(* IEC 61131-3 sources: test/Network/Pump, 1 file *)

(* ---- ONE_Pump_Table.st ---- *)
#define OBJECTS_CONFIG

//Define part of class pumpControl
#define test 1

FUNCTION GLOBAL TAB ONE_Pump
-1$UINT, 0$UINT,
0$UINT, 0$UINT,

1$UDINT,
TO_UDINT(2030910333), "pumpControl", 0$UINT, 0$UINT, 2$UINT,

_NO_ATTR, TO_UDINT(2903633677), "PUMPCONTROL1",
_NO_ATTR, TO_UDINT(874036919), "PUMPCONTROL2",

//Internal connections
0$UDINT,
0$UDINT,
0$UDINT,
0$UDINT,

//Initialization values
0$UDINT,
6$UDINT,
TO_UDINT(0), "MaxBorder", TO_UDINT(800),//|Pump.pumpControl1.MaxBorder;
TO_UDINT(0), "Pump", TO_UDINT(0),//|Pump.pumpControl1.Pump;
TO_UDINT(0), "ActFillLevel", TO_UDINT(0),//|Pump.pumpControl1.ActFillLevel;
TO_UDINT(1), "MaxBorder", TO_UDINT(800),//|Pump.pumpControl2.MaxBorder;
TO_UDINT(1), "Pump", TO_UDINT(0),//|Pump.pumpControl2.Pump;
TO_UDINT(1), "ActFillLevel", TO_UDINT(0),//|Pump.pumpControl2.ActFillLevel;

//Symbolic initialization values
0$UDINT,
0$UDINT,

//Initialization of string values
0$UDINT,
0$UDINT,

//Configuration of tasks (RealTime, Cyclic, Background)
0$UDINT,
0$UDINT,

0$UDINT,
2$UDINT,
TO_UDINT(0), (10)$UDINT, 4194303$DINT, 	//PUMPCONTROL1
TO_UDINT(1), (10)$UDINT, 4194303$DINT, 	//PUMPCONTROL2

0$UDINT,
0$UDINT,

//External connections
0$UDINT,
3$UDINT,
TO_UDINT(0), "ActFillLevel", C_TRY, TO_UDINT(1457099445), "AI0431","AI2",
TO_UDINT(0), "test2", C_TRY, TO_UDINT(4130059223), "SDM0811","Safe_Input1",
TO_UDINT(0), "test1", C_TRY, TO_UDINT(4130059223), "SDM0811","Safe_Input2",

//Magic internal connections
0$UDINT,
0$UDINT,

//Configuration of timeslots of tasks (RealTime, Cyclic)
#ifdef __LSLLDR_TIMESLOTS__
0$UDINT,
0$UDINT,

0$UDINT,
0$UDINT,

#endif //__LSLLDR_TIMESLOTS__

//MultiMaster connections
#ifdef __LSLLDR_MULTIMASTER__
0$UDINT,
0$UDINT,
#endif //__LSLLDR_MULTIMASTER__

//Configuration for task ID (RealTime, CyclicTime)
#ifdef __LSLLDR_TASKID__
"\\\\TASKS2  "
0$UDINT,
0$UDINT,

0$UDINT,
2$UDINT,
(0)$UDINT, 	//PUMPCONTROL1
(0)$UDINT, 	//PUMPCONTROL2

0$UDINT,
0$UDINT,

#endif //__LSLLDR_TASKID__

END_FUNCTION
